Fanuc KAREL source: KO00131.KL

PROGRAM KO00131
%NOLOCKGROUP
VAR
  R: REAL
  CFG: CONFIG
  OUT: XYZWPR
  N: ARRAY[2] OF BYTE
BEGIN
  N[1] = 1
  R = 2.0
  CFG.CFG_FLIP = TRUE
  OUT = POS(N[1], R, R, R, R, R, CFG)
END KO00131
